// TIA Portal V20 export
Screen "PN_DIAGNOSTIC ETH P4P5P6"  1276x673
  ScreenItem "Line_Header_X0_Y64" at 0,64 size 1276x0  Type=HmiLine
  ScreenItem "Title_ScreenOverview_X390_Y2" at 390,2 size 500x30  Type=HmiTextBox
  ScreenItem "PN-Diag_Reset" at 93,2 size 90x60  Type=HmiButton
  ScreenItem "PN-Diag_ReadNew" at 184,2 size 90x60  Type=HmiButton
  ScreenItem "Textfeld_1" at 292,8 size 95x22  Type=HmiTextBox
  ScreenItem "LED_1_Left_2" at 0,0 size 100x30  Type=HmiCircle
  ScreenItem "LED_1_Left_1" at 0,0 size 100x30  Type=HmiCircle
  ScreenItem "Textfeld_4" at 292,35 size 95x22  Type=HmiTextBox
  ScreenItem "permanentareaborderrectangle" at 0,0 size 0x0  Type=HmiRectangle
  ScreenItem "Button_Back" at 2,2 size 90x60  Type=HmiButton
  ScreenItem "PN-Diag_Counters" at 1093,2 size 90x60  Type=HmiButton
  ScreenItem "PN-Diag_LegendᆉY2" at 1184,2 size 90x60  Type=HmiButton
  ScreenItem "Rectangle_1" at 51,92 size 203x123  Type=HmiRectangle
  ScreenItem "LSicar_DeviceDiag_7" at 485,101 size 170x97  Type=HmiFaceplateContainer
  ScreenItem "LSicar_DeviceDiag_8" at 2294,628 size 170x97  Type=HmiFaceplateContainer
  ScreenItem "LSicar_DeviceDiag_9" at 293,277 size 170x97  Type=HmiFaceplateContainer
  ScreenItem "LSicar_DeviceDiag_2" at 1579,619 size 171x97  Type=HmiFaceplateContainer
  ScreenItem "LSicar_DeviceDiag_4" at 81,101 size 170x97  Type=HmiFaceplateContainer
  ScreenItem "LSicar_DeviceDiag_11" at 293,101 size 170x105  Type=HmiFaceplateContainer
  ScreenItem "LSicar_DeviceDiag_3" at 1942,495 size 170x97  Type=HmiFaceplateContainer
  ScreenItem "LSicar_DeviceDiag_5" at 2086,628 size 170x97  Type=HmiFaceplateContainer
  ScreenItem "LSicar_DeviceDiag_10" at 1604,81 size 170x97  Type=HmiFaceplateContainer
  ScreenItem "LSicar_DeviceDiag_12" at 680,446 size 170x97  Type=HmiFaceplateContainer
  ScreenItem "LSicar_DeviceDiag_1" at 485,277 size 170x97  Type=HmiFaceplateContainer
  ScreenItem "LSicar_DeviceDiag_6" at 2123,495 size 170x97  Type=HmiFaceplateContainer
  ScreenItem "LSicar_DeviceDiag_16" at 1375,728 size 170x97  Type=HmiFaceplateContainer
  ScreenItem "Faceplate container_1" at 880,104 size 170x100  Type=HmiFaceplateContainer
  ScreenItem "LSicar_DeviceDiag_13" at 2023,203 size 170x97  Type=HmiFaceplateContainer
  ScreenItem "线_4" at 190,162 size 60x0  Type=HmiLine
  ScreenItem "线_6" at 253,143 size 0x19  Type=HmiLine
  ScreenItem "线_26" at 254,142 size 129x0  Type=HmiLine
  ScreenItem "LSicar_DeviceDiag_17" at 61,269 size 170x105  Type=HmiFaceplateContainer
  ScreenItem "LSicar_DeviceDiag_18" at 680,101 size 170x97  Type=HmiFaceplateContainer
  ScreenItem "线_1" at 156,162 size 0x145  Type=HmiLine
  ScreenItem "线_3" at 363,152 size 23x0  Type=HmiLine
  ScreenItem "线_5" at 156,162 size 20x0  Type=HmiLine
  ScreenItem "线_7" at 363,153 size 0x54  Type=HmiLine
  ScreenItem "线_8" at 363,207 size 220x0  Type=HmiLine
  ScreenItem "线_9" at 583,179 size 0x27  Type=HmiLine
  ScreenItem "线_10" at 376,163 size 14x0  Type=HmiLine
  ScreenItem "线_11" at 376,163 size 0x54  Type=HmiLine
  ScreenItem "线_12" at 376,217 size 402x0  Type=HmiLine
  ScreenItem "线_13" at 778,179 size 0x37  Type=HmiLine
  ScreenItem "LSicar_DeviceDiag_19" at 293,446 size 170x97  Type=HmiFaceplateContainer
  ScreenItem "LSicar_DeviceDiag_20" at 1760,371 size 170x97  Type=HmiFaceplateContainer
  ScreenItem "LSicar_DeviceDiag_21" at 1941,371 size 170x97  Type=HmiFaceplateContainer
  ScreenItem "LSicar_DeviceDiag_22" at 2123,371 size 170x97  Type=HmiFaceplateContainer
  ScreenItem "LSicar_DeviceDiag_23" at 2309,371 size 170x97  Type=HmiFaceplateContainer
  ScreenItem "LSicar_DeviceDiag_24" at 1579,495 size 170x97  Type=HmiFaceplateContainer
  ScreenItem "LSicar_DeviceDiag_25" at 1760,495 size 170x97  Type=HmiFaceplateContainer
  ScreenItem "LSicar_DeviceDiag_26" at 1802,607 size 171x97  Type=HmiFaceplateContainer
  ScreenItem "Faceplate container_2" at 2309,495 size 170x97  Type=HmiFaceplateContainer
  ScreenItem "线_2" at 136,310 size 37x0  Type=HmiLine
  ScreenItem "线_14" at 136,310 size 0x79  Type=HmiLine
  ScreenItem "线_15" at 399,354 size 0x36  Type=HmiLine
  ScreenItem "线_16" at 411,354 size 0x36  Type=HmiLine
  ScreenItem "线_17" at 591,354 size 0x36  Type=HmiLine
  ScreenItem "线_24" at 136,390 size 262x0  Type=HmiLine
  ScreenItem "线_25" at 411,390 size 180x0  Type=HmiLine
  ScreenItem "线_29" at 120,320 size 52x0  Type=HmiLine
  ScreenItem "线_30" at 120,320 size 0x184  Type=HmiLine
  ScreenItem "线_31" at 375,514 size 0x43  Type=HmiLine
  ScreenItem "线_35" at 375,559 size 180x0  Type=HmiLine
  ScreenItem "线_36" at 120,503 size 282x0  Type=HmiLine
  ScreenItem "线_18" at 375,514 size 28x0  Type=HmiLine
  ScreenItem "LSicar_DeviceDiag_14" at 485,446 size 170x97  Type=HmiFaceplateContainer
  ScreenItem "线_33" at 566,516 size 0x43  Type=HmiLine
  ScreenItem "线_19" at 555,503 size 0x55  Type=HmiLine
  ScreenItem "线_20" at 555,503 size 39x0  Type=HmiLine
  ScreenItem "线_21" at 566,514 size 28x0  Type=HmiLine
  ScreenItem "LSicar_DeviceDiag_15" at 880,446 size 170x97  Type=HmiFaceplateContainer
  ScreenItem "线_22" at 566,559 size 233x0  Type=HmiLine
  ScreenItem "线_27" at 799,524 size 0x36  Type=HmiLine
  ScreenItem "线_28" at 811,523 size 0x36  Type=HmiLine
  ScreenItem "线_32" at 811,559 size 188x0  Type=HmiLine
  ScreenItem "线_34" at 999,523 size 0x36  Type=HmiLine
